Staubli VAL3: getTrajSize.pgx

public program getTrajSize(num& x_nSize)
begin
  x_nSize=size(trajTemp:tTrajItem)
end
